(* IEC 61131-3 sources: codesys-api/examples/mqtt_large_payload/st/probe, 2 files *)

(* ---- OnlineChangeProbe.st ---- *)
PROGRAM OnlineChangeProbe
// online_change_test.py rewrites this implementation in the session project and logs in with an online change;
// ProbeValue then shows that the new code runs. It does not touch the MQTT client.
VAR
	ProbeValue : UDINT;
END_VAR
// ---- implementation ----
ProbeValue := 0;

(* ---- UrlProbe.st ---- *)
PROGRAM UrlProbe
// The library's broker URL parsing (MQTT.STRING_TO_URL, as MQTT_CONTROL uses it) on a string written online:
// url_test.py checks user, password, host and port for credentials with '@', ':' and long passwords.
VAR
	Input : STRING(250);                    // written online; empty = idle
	Parsed : MQTT.URL;
	User : STRING(128);
	Password : STRING(128);
	Domain : STRING(80);
	Port : WORD;
	ParseCount : UDINT;
	LastInput : STRING(250);
END_VAR
// ---- implementation ----
IF Input <> '' AND Input <> LastInput THEN
	LastInput := Input;
	Parsed := MQTT.STRING_TO_URL(STR := Input, DEFAULT_PROTOCOL := '', DEFAULT_PATH := '/');
	User := Parsed.USER;
	Password := Parsed.PASSWORD;
	Domain := Parsed.DOMAIN;
	Port := Parsed.PORT;
	ParseCount := ParseCount + 1;
END_IF
